(* IEC 61131-3 sources: codesys-pass-demo/codesys/src, 11 files *)

(* ---- E_PassMode.st ---- *)
(*
 * E_PassMode
 * 目的 : PRG_Bench で、どの渡し方を測るかを選ぶ
 * 履歴 : 2026-11-03 新規作成
 *)
{attribute 'qualified_only'}  // CODESYS 拡張
{attribute 'strict'}          // CODESYS 拡張
TYPE E_PassMode :
(
    NONE     := 0,   (* 何もしない（基準の周期を見る） *)
    BY_INPUT := 1,   (* VAR_INPUT（コピー） *)
    BY_INOUT := 2,   (* VAR_IN_OUT CONSTANT（場所を渡す） *)
    BY_REF   := 3    (* REFERENCE TO（場所を登録） *)
);
END_TYPE

(* ---- ST_PassData.st ---- *)
(*
 * ST_PassData
 * 目的 : 渡し方の比較に使う構造体。
 *        小さいメンバー（モニタで見る用）と、大きい配列（コピーの重さを見る用）を持つ。
 * 履歴 : 2026-11-03 新規作成
 *)
TYPE ST_PassData :
STRUCT
    nCounter : DINT;    (* 毎サイクル更新。FB がどの値を見たかの目印 *)
    rValue   : REAL;    (* FB_ByInOutRW が書き換える *)
    bFlag    : BOOL;    (* 0.5 秒ごとに点滅。モニタで「生きている」のが見える *)
    aBig     : ARRAY[0..GVL_PassConst.N_BIG] OF DINT;   (* 16 KB。コピーの負荷を見る用 *)
END_STRUCT
END_TYPE

(* ---- GVL_PassConst.st ---- *)
(*
 * GVL_PassConst
 * 目的 : 確認用の定数
 * 履歴 : 2026-11-03 新規作成
 *)
{attribute 'qualified_only'}  // CODESYS 拡張: GVL_PassConst.N_BIG の形でしか書けなくする
VAR_GLOBAL CONSTANT
    N_BIG      : INT := 4095;   (* 大きい配列の上限。DINT × 4096 = 16 KB *)
    MAX_CALLS  : INT := 1000;   (* ベンチマークで1サイクルに呼ぶ回数の上限 *)
END_VAR

(* ---- GVL_PassTest.st ---- *)
(*
 * GVL_PassTest
 * 目的 : 3 つの FB に渡す「元データ」。全員がこれを見る。
 * 履歴 : 2026-11-03 新規作成
 *)
{attribute 'qualified_only'}  // CODESYS 拡張
VAR_GLOBAL
    stData : ST_PassData;
END_VAR

(* ---- FC_DisturbOtherTask.st ---- *)
(*
 * FC_DisturbOtherTask
 * 目的 : 「FB の処理の途中で、別のタスクが元データを書き換えた」状況を再現する。
 *        本物の別タスクだとタイミングが運任せになるので、FB の中からわざと呼んで必ず起こす。
 *        ※ 学習用。通常のコードで、FB の中から GVL を書き換えてはいけない。
 * 履歴 : 2026-11-03 新規作成
 *)
FUNCTION FC_DisturbOtherTask : BOOL
VAR CONSTANT
    N_JUMP : DINT := 1000;   (* 書き換えたことが一目で分かるよう、大きく足す *)
END_VAR

GVL_PassTest.stData.nCounter := GVL_PassTest.stData.nCounter + N_JUMP;
FC_DisturbOtherTask := TRUE;

(* ---- FB_ByInOutConst.st ---- *)
(*
 * FB_ByInOutConst
 * 目的 : VAR_IN_OUT CONSTANT（場所を渡す・読むだけ）の確認。
 *        コピーはせず、呼び出し元の変数そのものを見る。
 *
 * 確かめること:
 *   - 途中で元データが書き換わると、FB の中の値も変わる（bSnapshotKept = FALSE）
 *   - FB の中から書き換えようとするとコンパイルエラー（CONSTANT の効果）
 *   - 外から fbInOut.stIn は覗けない。モニタでどう表示されるか
 *
 * 入力 : stIn      呼び出し元のデータ（参照・読み取り専用）
 *        bDisturb  TRUE で、処理の途中に元データを書き換える
 * 出力 : FB_ByInput と同じ
 * 履歴 : 2026-11-03 新規作成
 *)
FUNCTION_BLOCK FB_ByInOutConst
VAR_IN_OUT CONSTANT
    stIn : ST_PassData;
END_VAR
VAR_INPUT
    bDisturb : BOOL;
END_VAR
VAR_OUTPUT
    nSeenFirst    : DINT;
    nSeenSecond   : DINT;
    bSnapshotKept : BOOL;
END_VAR

nSeenFirst := stIn.nCounter;
IF bDisturb THEN
    FC_DisturbOtherTask();
END_IF
nSeenSecond := stIn.nCounter;      // 元データを直接見ているので、+1000 された値が見える
bSnapshotKept := nSeenFirst = nSeenSecond;

// 実験: 下のコメントを外すとコンパイルエラー（CONSTANT なので書けない）
// stIn.nCounter := 0;

(* ---- FB_ByInOutRW.st ---- *)
(*
 * FB_ByInOutRW
 * 目的 : CONSTANT を付けない VAR_IN_OUT の確認（比較用・悪い例）。
 *        FB が呼び出し元の変数を書き換えられてしまう。
 *
 * 確かめること:
 *   - GVL_PassTest.stData.rValue が、この FB を呼ぶたびに +1 される
 *   - 「入力のつもりで渡したら、中身を変えられていた」が起きる
 *
 * 入出力 : stData  呼び出し元のデータ（参照・読み書き可）
 * 履歴 : 2026-11-03 新規作成
 *)
FUNCTION_BLOCK FB_ByInOutRW
VAR_IN_OUT
    stData : ST_PassData;
END_VAR

stData.rValue := stData.rValue + 1.0;   // 呼び出し元の rValue が書き換わる

(* ---- FB_ByInput.st ---- *)
(*
 * FB_ByInput
 * 目的 : VAR_INPUT（コピー渡し）の確認。
 *        呼んだ瞬間に構造体まるごとが FB の中へコピーされる。
 *
 * 確かめること:
 *   - 途中で元データが書き換わっても、FB の中の値は変わらない（bSnapshotKept = TRUE）
 *   - 外から fbInput.stIn を覗ける（モニタで展開できる）
 *
 * 入力 : stIn      渡されたデータ（コピー）
 *        bDisturb  TRUE で、処理の途中に元データを書き換える（別タスクの割り込みを再現）
 * 出力 : nSeenFirst / nSeenSecond  書き換え前後に FB が見た nCounter
 *        bSnapshotKept             前後で同じ値だったか
 * 履歴 : 2026-11-03 新規作成
 *)
FUNCTION_BLOCK FB_ByInput
VAR_INPUT
    stIn     : ST_PassData;
    bDisturb : BOOL;
END_VAR
VAR_OUTPUT
    nSeenFirst    : DINT;
    nSeenSecond   : DINT;
    bSnapshotKept : BOOL;
END_VAR

nSeenFirst := stIn.nCounter;
IF bDisturb THEN
    FC_DisturbOtherTask();          // 元データ（GVL）の nCounter を +1000
END_IF
nSeenSecond := stIn.nCounter;      // コピーなので、さっきと同じ値のはず
bSnapshotKept := nSeenFirst = nSeenSecond;

// 実験: 下のコメントを外してもコンパイルは通る。書き換わるのは FB 内のコピーだけで、元データは無傷
// stIn.nCounter := 0;

(* ---- FB_ByRef.st ---- *)
(*
 * FB_ByRef
 * 目的 : REFERENCE TO（場所を登録しておく）の確認。CODESYS 独自の機能。
 *        呼び出し側が  fbRef.refIn REF= 変数;  で場所を登録してから呼ぶ。
 *
 * 確かめること:
 *   - VAR_IN_OUT と同じく、途中の書き換えが見える（bSnapshotKept = FALSE）
 *   - 登録していないインスタンスは bRefValid = FALSE になり、何もしない
 *   - 外から fbRef.refIn を覗いたとき、モニタでどう表示されるか
 *
 * 入力 : refIn     データの場所（REF= で登録）
 *        bDisturb  TRUE で、処理の途中に元データを書き換える
 * 出力 : bRefValid  refIn が有効か（__ISVALIDREF の結果）
 *        ほかは FB_ByInput と同じ
 * 履歴 : 2026-11-03 新規作成
 *)
FUNCTION_BLOCK FB_ByRef
VAR_INPUT
    refIn    : REFERENCE TO ST_PassData;   // CODESYS 拡張（IEC 61131-3 の標準ではない）
    bDisturb : BOOL;
END_VAR
VAR_OUTPUT
    bRefValid     : BOOL;
    nSeenFirst    : DINT;
    nSeenSecond   : DINT;
    bSnapshotKept : BOOL;
END_VAR

// 登録されていない参照を読むと例外で PLC が止まる。必ず先に確かめる
bRefValid := __ISVALIDREF(refIn);   // CODESYS 拡張
IF NOT bRefValid THEN
    nSeenFirst    := 0;
    nSeenSecond   := 0;
    bSnapshotKept := FALSE;
    RETURN;
END_IF

nSeenFirst := refIn.nCounter;      // 普通の変数と同じ書き方で読める
IF bDisturb THEN
    FC_DisturbOtherTask();
END_IF
nSeenSecond := refIn.nCounter;
bSnapshotKept := nSeenFirst = nSeenSecond;

// 実験: 下のコメントを外すとコンパイルは通り、元データが書き換わる（REFERENCE には CONSTANT がない）
// refIn.nCounter := 0;

(* ---- PRG_Bench.st ---- *)
(*
 * PRG_Bench
 * 目的 : 渡し方による処理時間の違いを見る。
 *        選んだ渡し方で、16 KB の構造体を nCalls 回 FB に渡す。
 *        BenchTask の周期時間を「タスク設定 → モニタ」で見て比べる。
 *
 * モニタから切り替えるもの:
 *   eMode   NONE / BY_INPUT / BY_INOUT / BY_REF
 *   nCalls  1 サイクルに呼ぶ回数（0〜MAX_CALLS）
 *
 * 履歴 : 2026-11-03 新規作成
 *)
PROGRAM PRG_Bench
VAR
    eMode    : E_PassMode := E_PassMode.NONE;
    nCalls   : INT := 100;
    nDone    : INT;           (* 実際に呼んだ回数 *)
    i        : INT;
    fbInput  : FB_ByInput;
    fbInOut  : FB_ByInOutConst;
    fbRef    : FB_ByRef;
END_VAR

nCalls := LIMIT(0, nCalls, GVL_PassConst.MAX_CALLS);   // ループ回数に上限を置く
nDone  := 0;

CASE eMode OF
E_PassMode.NONE:
    ;   // 何もしない。この時の周期時間が基準

E_PassMode.BY_INPUT:
    FOR i := 1 TO nCalls DO
        fbInput(stIn := GVL_PassTest.stData, bDisturb := FALSE);   // 毎回 16 KB コピー
        nDone := nDone + 1;
    END_FOR

E_PassMode.BY_INOUT:
    FOR i := 1 TO nCalls DO
        fbInOut(stIn := GVL_PassTest.stData, bDisturb := FALSE);   // 場所だけ渡す
        nDone := nDone + 1;
    END_FOR

E_PassMode.BY_REF:
    fbRef.refIn REF= GVL_PassTest.stData;                         // CODESYS 拡張
    FOR i := 1 TO nCalls DO
        fbRef(bDisturb := FALSE);
        nDone := nDone + 1;
    END_FOR

ELSE
    eMode := E_PassMode.NONE;
END_CASE

(* ---- PRG_PassDemo.st ---- *)
(*
 * PRG_PassDemo
 * 目的 : 3 つの渡し方を、同じ元データ・同じ条件で並べて呼ぶ。
 *        オンラインでこの PRG を開き、各インスタンスを展開して見比べる。
 *
 * モニタから切り替えるもの（書き込み値を入れて Ctrl+F7）:
 *   bDisturb        TRUE: FB の処理途中で元データを書き換える
 *   bRefEveryCycle  TRUE: 毎サイクル REF= し直す / FALSE: 最初の1回だけ
 *
 * 履歴 : 2026-11-03 新規作成
 *)
PROGRAM PRG_PassDemo
VAR
    fbInput        : FB_ByInput;
    fbInOut        : FB_ByInOutConst;
    fbRef          : FB_ByRef;
    fbRefNotLinked : FB_ByRef;          (* わざと REF= しない。bRefValid = FALSE になるのを見る *)
    fbInOutRW      : FB_ByInOutRW;

    nCycle         : DINT;
    bDisturb       : BOOL := TRUE;
    bRefEveryCycle : BOOL := TRUE;
    bRefLinked     : BOOL;
    tonBlink       : TON;

    nDataSize      : UDINT;             (* 構造体の大きさ [byte]。コピーされる量の目安 *)
    nInstSizeInput : UDINT;             (* FB インスタンスの大きさ [byte] *)
    nInstSizeInOut : UDINT;
    nInstSizeRef   : UDINT;
END_VAR
VAR CONSTANT
    T_BLINK : TIME := T#500MS;
END_VAR

nCycle := nCycle + 1;

(* 元データを毎サイクル作り直す。FB ごとの比較を同じ条件にするため *)
tonBlink(IN := NOT tonBlink.Q, PT := T_BLINK);
IF tonBlink.Q THEN
    GVL_PassTest.stData.bFlag := NOT GVL_PassTest.stData.bFlag;
END_IF
GVL_PassTest.stData.aBig[0]                   := nCycle;
GVL_PassTest.stData.aBig[GVL_PassConst.N_BIG] := -nCycle;

(* ---- 1. VAR_INPUT（コピー） ---- *)
GVL_PassTest.stData.nCounter := nCycle;
fbInput(stIn := GVL_PassTest.stData, bDisturb := bDisturb);

(* ---- 2. VAR_IN_OUT CONSTANT（場所を渡す） ---- *)
GVL_PassTest.stData.nCounter := nCycle;          // 1. で +1000 された分を戻す
fbInOut(stIn := GVL_PassTest.stData, bDisturb := bDisturb);

(* ---- 3. REFERENCE TO（場所を登録） ---- *)
GVL_PassTest.stData.nCounter := nCycle;
IF bRefEveryCycle OR NOT bRefLinked THEN
    fbRef.refIn REF= GVL_PassTest.stData;        // CODESYS 拡張
    bRefLinked := TRUE;
END_IF
fbRef(bDisturb := bDisturb);

fbRefNotLinked(bDisturb := FALSE);              // refIn 未登録のまま呼ぶ

(* ---- 4. CONSTANT なしの VAR_IN_OUT（比較用） ---- *)
fbInOutRW(stData := GVL_PassTest.stData);       // stData.rValue が毎サイクル +1 される

(* 最後に、元データの nCounter を正しい値に戻しておく *)
GVL_PassTest.stData.nCounter := nCycle;

(* 大きさの確認 *)
nDataSize      := SIZEOF(GVL_PassTest.stData);
nInstSizeInput := SIZEOF(fbInput);    // 16 KB 超のはず（コピーを中に持つ）
nInstSizeInOut := SIZEOF(fbInOut);    // 小さいはず（場所だけ持つ）
nInstSizeRef   := SIZEOF(fbRef);      // 小さいはず（場所だけ持つ）

(* ---- 実験：1行ずつコメントを外して、コンパイル結果を見る ----
   nCycle := fbInOut.stIn.nCounter;   // VAR_IN_OUT は外から読めない → エラーの予想
   fbInOut(bDisturb := FALSE);        // VAR_IN_OUT を渡さずに呼ぶ → エラーの予想
   nCycle := fbRef.refIn.nCounter;    // REFERENCE は外から読める → 通る予想
   nCycle := fbInput.stIn.nCounter;   // VAR_INPUT は外から読める → 通る予想
*)
